Fanuc KAREL source: kd00031.KL

-- PROVISIONAL review KL for V770-1; original PC SHA256 4364f114a299508c982d9f5eda2ab294f865ac170deacf7f63ef5bfcb9fb63a2
-- Incomplete behavior may be omitted. Consult companion uncertainty JSON. Do not deploy.
PROGRAM KD00031
%NOLOCKGROUP
VAR
  I : INTEGER
  J : INTEGER
  B : BOOLEAN
  R : REAL
  S : STRING[80]
BEGIN
  -- UNRESOLVED_PC offsets 5-21; opcodes 9D,81,18,9C,12,22,9D,13,04
  -- UNRESOLVED_PC offsets 26-30; opcodes 7F
END KD00031
